(* PLC project Vn_ld_two_coils, Beckhoff Automation GmbH TwinCAT PLC Control 3.5.13.21 *)
(* stored: creationDateTime 1970-01-01T00:00:00 *)

PROGRAM Vn_ld_two_coils

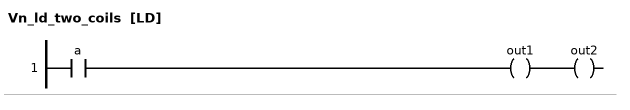
(* LD diagram, written out as Structured Text *)
out1 := a;
out2 := a;
END_PROGRAM
